// TIA Portal V20 export
// export: Created 2026-10-20T12:51:26.8635098Z, ExportSetting WithDefaults, DisplayName Totally Integrated Automation Portal, DisplayVersion V20 Update 6, DisplayName TIA Portal Openness, DisplayVersion V20 Update 6, DisplayName TIA Portal Version Control Interface, DisplayVersion V20 Update 6, DisplayName SINAMICS Startdrive Advanced, DisplayVersion V20 SP1, DisplayName SINAMICS Startdrive G130, G150, S120, S150, SINAMICS MV, G220, S200, S210, DisplayVersion V20 SP1, DisplayName SINAMICS Startdrive G110M, G120, G120C, G120D, G120P, G115D, DisplayVersion V20 SP1, DisplayName STEP 7 Professional, DisplayVersion V20 Update 6, DisplayName STEP 7 Safety, DisplayVersion V20 Update 2, DisplayName WinCC Basic/Comfort/Advanced, DisplayVersion V20 Update 6, DisplayName WinCC Unified, DisplayVersion V20 Update 6
FUNCTION "Overhang_IO_FC" : Void   // FC40, F_LAD
{ S7_Optimized_Access := 'TRUE' }
VERSION : 0.1
// stored: AutoNumber true, IsIECCheckEnabled false, UDAEnableTagReadback false
BEGIN

REGION Network 1: SYSTEM 1
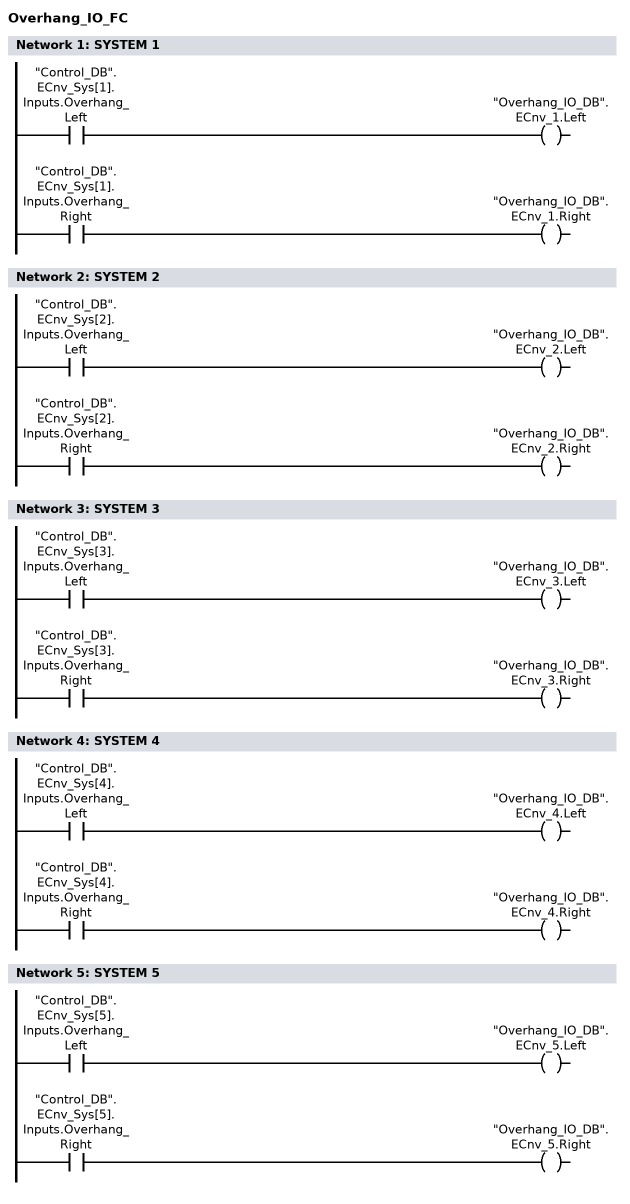
   RUNG wire#powerrail
      Contact( "Control_DB".ECnv_Sys[1].Inputs.Overhang_Left )
      Coil( "Overhang_IO_DB".ECnv_1.Left )
   END_RUNG
   RUNG wire#powerrail
      Contact( "Control_DB".ECnv_Sys[1].Inputs.Overhang_Right )
      Coil( "Overhang_IO_DB".ECnv_1.Right )
   END_RUNG
   // the same network as SCL:
   "Overhang_IO_DB".ECnv_1.Left := "Control_DB".ECnv_Sys[1].Inputs.Overhang_Left;
   "Overhang_IO_DB".ECnv_1.Right := "Control_DB".ECnv_Sys[1].Inputs.Overhang_Right;
END_REGION

REGION Network 2: SYSTEM 2
   RUNG wire#powerrail
      Contact( "Control_DB".ECnv_Sys[2].Inputs.Overhang_Left )
      Coil( "Overhang_IO_DB".ECnv_2.Left )
   END_RUNG
   RUNG wire#powerrail
      Contact( "Control_DB".ECnv_Sys[2].Inputs.Overhang_Right )
      Coil( "Overhang_IO_DB".ECnv_2.Right )
   END_RUNG
   // the same network as SCL:
   "Overhang_IO_DB".ECnv_2.Left := "Control_DB".ECnv_Sys[2].Inputs.Overhang_Left;
   "Overhang_IO_DB".ECnv_2.Right := "Control_DB".ECnv_Sys[2].Inputs.Overhang_Right;
END_REGION

REGION Network 3: SYSTEM 3
   RUNG wire#powerrail
      Contact( "Control_DB".ECnv_Sys[3].Inputs.Overhang_Left )
      Coil( "Overhang_IO_DB".ECnv_3.Left )
   END_RUNG
   RUNG wire#powerrail
      Contact( "Control_DB".ECnv_Sys[3].Inputs.Overhang_Right )
      Coil( "Overhang_IO_DB".ECnv_3.Right )
   END_RUNG
   // the same network as SCL:
   "Overhang_IO_DB".ECnv_3.Left := "Control_DB".ECnv_Sys[3].Inputs.Overhang_Left;
   "Overhang_IO_DB".ECnv_3.Right := "Control_DB".ECnv_Sys[3].Inputs.Overhang_Right;
END_REGION

REGION Network 4: SYSTEM 4
   RUNG wire#powerrail
      Contact( "Control_DB".ECnv_Sys[4].Inputs.Overhang_Left )
      Coil( "Overhang_IO_DB".ECnv_4.Left )
   END_RUNG
   RUNG wire#powerrail
      Contact( "Control_DB".ECnv_Sys[4].Inputs.Overhang_Right )
      Coil( "Overhang_IO_DB".ECnv_4.Right )
   END_RUNG
   // the same network as SCL:
   "Overhang_IO_DB".ECnv_4.Left := "Control_DB".ECnv_Sys[4].Inputs.Overhang_Left;
   "Overhang_IO_DB".ECnv_4.Right := "Control_DB".ECnv_Sys[4].Inputs.Overhang_Right;
END_REGION

REGION Network 5: SYSTEM 5
   RUNG wire#powerrail
      Contact( "Control_DB".ECnv_Sys[5].Inputs.Overhang_Left )
      Coil( "Overhang_IO_DB".ECnv_5.Left )
   END_RUNG
   RUNG wire#powerrail
      Contact( "Control_DB".ECnv_Sys[5].Inputs.Overhang_Right )
      Coil( "Overhang_IO_DB".ECnv_5.Right )
   END_RUNG
   // the same network as SCL:
   "Overhang_IO_DB".ECnv_5.Left := "Control_DB".ECnv_Sys[5].Inputs.Overhang_Left;
   "Overhang_IO_DB".ECnv_5.Right := "Control_DB".ECnv_Sys[5].Inputs.Overhang_Right;
END_REGION
END_FUNCTION
